  MoveL 497 to (87.59, -0.5, 58.1) mm, rotated rx 0 ry 90 rz 0 deg; joints [-13.797, -57.781, 117.086, 164.062, 60.282, -81.942]
  MoveL 498 to (93.3, -5.75, 58.1) mm, rotated rx 0 ry 90 rz 0 deg; joints [-13.739, -57.804, 116.577, 164.043, 59.762, -81.806]
  MoveL 499 to (99.9, -9.83, 58.1) mm, rotated rx 0 ry 90 rz 0 deg; joints [-13.673, -57.72, 116.001, 164.04, 59.279, -81.688]
  MoveL 500 to (107.03, -12.94, 58.1) mm, rotated rx 0 ry 90 rz 0 deg; joints [-13.603, -57.557, 115.386, 164.047, 58.834, -81.585]
  MoveL 501 to (114.36, -15.46, 58.1) mm, rotated rx 0 ry 90 rz 0 deg; joints [-13.531, -57.352, 114.755, 164.059, 58.415, -81.491]
  MoveL 502 to (121.65, -18.1, 58.1) mm, rotated rx 0 ry 90 rz 0 deg; joints [-13.46, -57.151, 114.125, 164.068, 57.991, -81.396]
  MoveL 503 to (126.38, -19.97, 58.1) mm, rotated rx 0 ry 90 rz 0 deg; joints [-13.414, -57.027, 113.713, 164.072, 57.707, -81.331]
  MoveL 504 to (131.09, -21.86, 58.1) mm, rotated rx 0 ry 90 rz 0 deg; joints [-13.369, -56.903, 113.3, 164.074, 57.422, -81.265]
  MoveL 505 to (135.76, -23.86, 58.1) mm, rotated rx 0 ry 90 rz 0 deg; joints [-13.325, -56.786, 112.889, 164.074, 57.133, -81.198]
  MoveL 506 to (140.36, -26.03, 58.1) mm, rotated rx 0 ry 90 rz 0 deg; joints [-13.281, -56.679, 112.48, 164.072, 56.837, -81.127]
  MoveL 507 to (145.03, -27.98, 58.1) mm, rotated rx 0 ry 90 rz 0 deg; joints [-13.237, -56.555, 112.066, 164.071, 56.55, -81.06]
  MoveL 508 to (150, -29.16, 58.1) mm, rotated rx 0 ry 90 rz 0 deg; joints [-13.191, -56.379, 111.633, 164.079, 56.296, -81.006]
  MoveL 509 to (150, -26.31, 58.1) mm, rotated rx 0 ry 90 rz 0 deg; joints [-13.191, -56.239, 111.66, 164.11, 56.456, -81.061]
  MoveL 510 to (146.2, -24.88, 58.1) mm, rotated rx 0 ry 90 rz 0 deg; joints [-13.226, -56.348, 111.996, 164.109, 56.681, -81.112]
  MoveL 511 to (142.73, -22.75, 58.1) mm, rotated rx 0 ry 90 rz 0 deg; joints [-13.259, -56.405, 112.31, 164.117, 56.932, -81.175]
  MoveL 512 to (139.28, -20.57, 58.1) mm, rotated rx 0 ry 90 rz 0 deg; joints [-13.291, -56.458, 112.622, 164.124, 57.187, -81.239]
  MoveL 513 to (135.74, -18.56, 58.1) mm, rotated rx 0 ry 90 rz 0 deg; joints [-13.325, -56.522, 112.938, 164.129, 57.434, -81.299]
  MoveL 514 to (132.21, -16.55, 58.1) mm, rotated rx 0 ry 90 rz 0 deg; joints [-13.358, -56.585, 113.253, 164.134, 57.682, -81.36]
  MoveL 515 to (127.82, -13.81, 58.1) mm, rotated rx 0 ry 90 rz 0 deg; joints [-13.4, -56.649, 113.645, 164.141, 58.004, -81.44]
  MoveL 516 to (123.5, -10.92, 58.1) mm, rotated rx 0 ry 90 rz 0 deg; joints [-13.442, -56.7, 114.031, 164.15, 58.332, -81.522]
  MoveL 517 to (119.33, -7.82, 58.1) mm, rotated rx 0 ry 90 rz 0 deg; joints [-13.482, -56.732, 114.405, 164.16, 58.666, -81.607]
  MoveL 518 to (115.6, -4.28, 58.1) mm, rotated rx 0 ry 90 rz 0 deg; joints [-13.518, -56.719, 114.744, 164.176, 59.011, -81.698]
  MoveL 519 to (112.62, 0, 58.1) mm, rotated rx 0 ry 90 rz 0 deg; joints [-13.548, -56.631, 115.024, 164.202, 59.369, -81.797]
  MoveL 520 to (-12.62, 0, 58.1) mm, rotated rx 0 ry 90 rz 0 deg; joints [-14.893, -62.159, 125.079, 163.369, 63.9, -82.514]
  MoveL 521 to (-15.6, -4.28, 58.1) mm, rotated rx 0 ry 90 rz 0 deg; joints [-14.928, -62.542, 125.276, 163.304, 63.726, -82.437]
  MoveL 522 to (-19.33, -7.82, 58.1) mm, rotated rx 0 ry 90 rz 0 deg; joints [-14.973, -62.916, 125.535, 163.239, 63.623, -82.379]
  MoveL 523 to (-23.5, -10.92, 58.1) mm, rotated rx 0 ry 90 rz 0 deg; joints [-15.023, -63.282, 125.831, 163.173, 63.561, -82.331]
  MoveL 524 to (-27.82, -13.81, 58.1) mm, rotated rx 0 ry 90 rz 0 deg; joints [-15.074, -63.645, 126.138, 163.108, 63.515, -82.287]
  MoveL 525 to (-32.2, -16.55, 58.1) mm, rotated rx 0 ry 90 rz 0 deg; joints [-15.128, -64.002, 126.45, 163.043, 63.478, -82.246]
  MoveL 526 to (-35.74, -18.56, 58.1) mm, rotated rx 0 ry 90 rz 0 deg; joints [-15.171, -64.279, 126.702, 162.991, 63.461, -82.217]
  MoveL 527 to (-39.28, -20.57, 58.1) mm, rotated rx 0 ry 90 rz 0 deg; joints [-15.214, -64.557, 126.953, 162.939, 63.442, -82.187]
  MoveL 528 to (-42.73, -22.75, 58.1) mm, rotated rx 0 ry 90 rz 0 deg; joints [-15.257, -64.841, 127.196, 162.886, 63.407, -82.152]
  MoveL 529 to (-46.2, -24.88, 58.1) mm, rotated rx 0 ry 90 rz 0 deg; joints [-15.3, -65.125, 127.439, 162.833, 63.375, -82.118]
  MoveL 530 to (-50, -26.31, 58.1) mm, rotated rx 0 ry 90 rz 0 deg; joints [-15.347, -65.381, 127.714, 162.783, 63.399, -82.1]
  MoveL 531 to (-50, -26.31, 103.1) mm, rotated rx 0 ry 90 rz 0 deg; joints [-17.375, -64.79, 126.71, 160.473, 63.306, -80.948]
  Sollgeschwindigkeit (200.0 mm/s)
  MoveL 532 to (-42.49, -26.16, 103.1) mm, rotated rx 0 ry 90 rz 0 deg; joints [-17.271, -64.448, 126.142, 160.55, 63.077, -80.915]
  MoveL 533 to (-34.99, -26.02, 103.1) mm, rotated rx 0 ry 90 rz 0 deg; joints [-17.168, -64.106, 125.572, 160.625, 62.845, -80.882]
  MoveL 534 to (-27.48, -25.87, 103.1) mm, rotated rx 0 ry 90 rz 0 deg; joints [-17.066, -63.763, 124.999, 160.699, 62.612, -80.848]
  MoveL 535 to (-19.97, -25.73, 103.1) mm, rotated rx 0 ry 90 rz 0 deg; joints [-16.966, -63.42, 124.425, 160.771, 62.377, -80.814]
  MoveL 536 to (-12.46, -25.58, 103.1) mm, rotated rx 0 ry 90 rz 0 deg; joints [-16.866, -63.077, 123.848, 160.842, 62.141, -80.778]
  MoveL 537 to (-4.96, -25.43, 103.1) mm, rotated rx 0 ry 90 rz 0 deg; joints [-16.768, -62.734, 123.268, 160.911, 61.902, -80.742]
  MoveL 538 to (2.55, -25.29, 103.1) mm, rotated rx 0 ry 90 rz 0 deg; joints [-16.671, -62.39, 122.687, 160.978, 61.661, -80.706]
  MoveL 539 to (10.05, -25.14, 103.1) mm, rotated rx 0 ry 90 rz 0 deg; joints [-16.575, -62.046, 122.103, 161.043, 61.419, -80.668]
  MoveL 540 to (17.56, -25, 103.1) mm, rotated rx 0 ry 90 rz 0 deg; joints [-16.48, -61.701, 121.516, 161.107, 61.175, -80.63]
  MoveL 541 to (25.07, -24.85, 103.1) mm, rotated rx 0 ry 90 rz 0 deg; joints [-16.386, -61.356, 120.927, 161.17, 60.929, -80.592]
  MoveL 542 to (32.58, -24.71, 103.1) mm, rotated rx 0 ry 90 rz 0 deg; joints [-16.293, -61.011, 120.336, 161.231, 60.681, -80.552]
  MoveL 543 to (40.08, -24.56, 103.1) mm, rotated rx 0 ry 90 rz 0 deg; joints [-16.201, -60.665, 119.742, 161.29, 60.431, -80.512]
  Sollgeschwindigkeit (50.0 mm/s)
  MoveL 544 to (40.08, -24.56, 58.1) mm, rotated rx 0 ry 90 rz 0 deg; joints [-14.296, -61.22, 120.719, 163.524, 60.538, -81.724]
  MoveL 545 to (36.66, -28.17, 58.1) mm, rotated rx 0 ry 90 rz 0 deg; joints [-14.334, -61.573, 120.955, 163.463, 60.432, -81.665]
  MoveL 546 to (36.08, -29.02, 58.1) mm, rotated rx 0 ry 90 rz 0 deg; joints [-14.34, -61.646, 120.993, 163.45, 60.399, -81.65]
  MoveL 547 to (35.49, -29.88, 58.1) mm, rotated rx 0 ry 90 rz 0 deg; joints [-14.346, -61.72, 121.031, 163.437, 60.366, -81.634]
  MoveL 548 to (34.9, -30.69, 58.08) mm, rotated rx 90 ry 86.96 rz 90 deg; joints [-14.257, -62.836, 120.907, 163.332, 59.164, -84.313]
  MoveL 549 to (34.32, -31.5, 58.01) mm, rotated rx 90 ry 83.41 rz 90 deg; joints [-14.096, -64.109, 120.741, 163.266, 57.761, -87.482]
  MoveL 550 to (33.73, -32.31, 57.9) mm, rotated rx 90 ry 79.85 rz 90 deg; joints [-13.873, -65.357, 120.562, 163.261, 56.359, -90.69]
  MoveL 551 to (33.17, -33.03, 57.74) mm, rotated rx 90 ry 76.63 rz 90 deg; joints [-13.62, -66.464, 120.392, 163.313, 55.094, -93.64]
  MoveL 552 to (32.6, -33.74, 57.55) mm, rotated rx 90 ry 73.4 rz 90 deg; joints [-13.318, -67.543, 120.214, 163.421, 53.837, -96.635]
  MoveL 553 to (32.04, -34.44, 57.32) mm, rotated rx 90 ry 70.18 rz 90 deg; joints [-12.968, -68.591, 120.028, 163.59, 52.593, -99.681]
  MoveL 554 to (31.48, -35.13, 57.05) mm, rotated rx 90 ry 66.95 rz 90 deg; joints [-12.57, -69.605, 119.836, 163.822, 51.364, -102.781]
  MoveL 555 to (30.63, -35.95, 56.67) mm, rotated rx 90 ry 63.01 rz 90 deg; joints [-12.022, -70.803, 119.607, 164.198, 49.895, -106.656]
  MoveL 556 to (29.79, -36.73, 56.24) mm, rotated rx 90 ry 59.07 rz 90 deg; joints [-11.405, -71.942, 119.374, 164.681, 48.463, -110.633]
  MoveL 557 to (28.94, -37.49, 55.75) mm, rotated rx 90 ry 55.13 rz 90 deg; joints [-10.723, -73.018, 119.14, 165.281, 47.076, -114.724]
  MoveL 558 to (28.04, -38.22, 55.2) mm, rotated rx 90 ry 51.13 rz 90 deg; joints [-9.964, -74.045, 118.907, 166.015, 45.723, -119.006]
  MoveL 559 to (27.13, -38.91, 54.6) mm, rotated rx 90 ry 47.13 rz 90 deg; joints [-9.143, -74.999, 118.678, 166.882, 44.436, -123.425]
  MoveL 560 to (26.62, -39.4, 54.13) mm, rotated rx 90 ry 44.19 rz 90 deg; joints [-8.5, -75.643, 118.503, 167.608, 43.534, -126.764]
  MoveL 561 to (26.11, -39.85, 53.64) mm, rotated rx 90 ry 41.24 rz 90 deg; joints [-7.827, -76.243, 118.333, 168.411, 42.677, -130.182]
  MoveL 562 to (25.61, -40.28, 53.12) mm, rotated rx 90 ry 38.3 rz 90 deg; joints [-7.124, -76.8, 118.17, 169.291, 41.869, -133.682]
  MoveL 563 to (25.48, -40.77, 52.46) mm, rotated rx 90 ry 34.73 rz 90 deg; joints [-6.232, -77.386, 117.944, 170.466, 40.951, -138.045]
  MoveL 564 to (25.37, -41.21, 51.78) mm, rotated rx 90 ry 31.15 rz 90 deg; joints [-5.304, -77.904, 117.731, 171.753, 40.121, -142.525]
  MoveL 565 to (25.25, -41.61, 51.06) mm, rotated rx 90 ry 27.57 rz 90 deg; joints [-4.344, -78.351, 117.534, 173.144, 39.385, -147.116]
  MoveL 566 to (25.45, -41.88, 50.53) mm, rotated rx 90 ry 24.95 rz 90 deg; joints [-3.621, -78.616, 117.379, 174.228, 38.905, -150.548]
  MoveL 567 to (25.65, -42.12, 49.98) mm, rotated rx 90 ry 22.33 rz 90 deg; joints [-2.886, -78.842, 117.233, 175.359, 38.482, -154.03]
  MoveL 568 to (26.42, -42.43, 49.12) mm, rotated rx 90 ry 18.35 rz 90 deg; joints [-1.747, -79.083, 116.996, 177.159, 37.948, -159.407]
  MoveL 569 to (27.19, -42.54, 48.79) mm, rotated rx 90 ry 16.83 rz 90 deg; joints [-1.304, -79.122, 116.877, 177.871, 37.774, -161.491]
  MoveL 570 to (27.95, -42.64, 48.46) mm, rotated rx 90 ry 15.3 rz 90 deg; joints [-0.86, -79.147, 116.761, 178.592, 37.622, -163.585]
  MoveL 571 to (28.72, -42.72, 48.12) mm, rotated rx 90 ry 13.77 rz 90 deg; joints [-0.413, -79.159, 116.649, 179.321, 37.492, -165.687]
  MoveL 572 to (29.56, -42.79, 47.84) mm, rotated rx 90 ry 12.53 rz 90 deg; joints [-0.048, -79.145, 116.544, 179.921, 37.398, -167.409]
  MoveL 573 to (30.4, -42.85, 47.56) mm, rotated rx 90 ry 11.28 rz 90 deg; joints [0.318, -79.123, 116.442, -179.476, 37.32, -169.135]
  MoveL 574 to (31.24, -42.9, 47.28) mm, rotated rx 90 ry 10.04 rz 90 deg; joints [0.684, -79.092, 116.342, -178.87, 37.256, -170.862]
  MoveL 575 to (31.96, -42.97, 46.87) mm, rotated rx 90 ry 8.2 rz 90 deg; joints [1.225, -79.061, 116.239, -177.974, 37.195, -173.413]
  MoveL 576 to (32.69, -43.02, 46.45) mm, rotated rx 90 ry 6.37 rz 90 deg; joints [1.765, -79.012, 116.143, -177.078, 37.167, -175.965]
  MoveL 577 to (33.42, -43.06, 46.03) mm, rotated rx 90 ry 4.53 rz 90 deg; joints [2.305, -78.943, 116.052, -176.183, 37.17, -178.514]
  MoveL 578 to (34.18, -43.09, 45.39) mm, rotated rx 90 ry 1.71 rz 90 deg; joints [3.132, -78.823, 115.951, -174.82, 37.241, 177.584]
  MoveL 579 to (34.94, -43.1, 44.73) mm, rotated rx 90 ry 0 rz 90 deg; joints [3.644, -78.708, 115.873, -173.982, 37.317, 175.208]
  MoveL 580 to (35.7, -43.1, 44.06) mm, rotated rx 90 ry 0 rz 90 deg; joints [3.672, -78.658, 115.812, -173.934, 37.308, 175.169]
  MoveL 581 to (37.13, -43.1, 42.71) mm, rotated rx 90 ry 0 rz 90 deg; joints [3.729, -78.564, 115.695, -173.837, 37.292, 175.09]
  MoveL 582 to (38.7, -43.1, 41.89) mm, rotated rx 90 ry 0 rz 90 deg; joints [3.762, -78.463, 115.572, -173.78, 37.272, 175.043]
  MoveL 583 to (40.05, -43.1, 41.81) mm, rotated rx 90 ry 0 rz 90 deg; joints [3.762, -78.378, 115.468, -173.778, 37.252, 175.04]
  MoveL 584 to (41.5, -43.1, 42.11) mm, rotated rx 90 ry 0 rz 90 deg; joints [3.744, -78.29, 115.359, -173.805, 37.231, 175.06]
  MoveL 585 to (45.39, -43.1, 43.71) mm, rotated rx 90 ry 0 rz 90 deg; joints [3.66, -78.055, 115.069, -173.934, 37.169, 175.16]
  MoveL 586 to (47.73, -43.1, 44.54) mm, rotated rx 90 ry 0 rz 90 deg; joints [3.616, -77.913, 114.892, -174.003, 37.131, 175.212]
  MoveL 587 to (50.09, -43.1, 44.8) mm, rotated rx 90 ry 0 rz 90 deg; joints [3.598, -77.767, 114.712, -174.028, 37.095, 175.23]
  MoveL 588 to (53.81, -43.1, 44.03) mm, rotated rx 90 ry 0 rz 90 deg; joints [3.621, -77.534, 114.421, -173.981, 37.04, 175.189]
  MoveL 589 to (56.17, -43.1, 43.02) mm, rotated rx 90 ry 0 rz 90 deg; joints [3.66, -77.383, 114.234, -173.912, 37.006, 175.132]
  MoveL 590 to (58.51, -43.1, 42.11) mm, rotated rx 90 ry 0 rz 90 deg; joints [3.694, -77.235, 114.049, -173.85, 36.972, 175.08]
  MoveL 591 to (60.69, -43.1, 41.79) mm, rotated rx 90 ry 0 rz 90 deg; joints [3.702, -77.099, 113.877, -173.832, 36.938, 175.064]
  MoveL 592 to (62.64, -43.1, 42.54) mm, rotated rx 90 ry 0 rz 90 deg; joints [3.663, -76.981, 113.73, -173.893, 36.905, 175.11]
  MoveL 593 to (64.38, -43.1, 44.14) mm, rotated rx 90 ry 0 rz 90 deg; joints [3.587, -76.88, 113.602, -174.015, 36.872, 175.206]
  MoveL 594 to (65.25, -43.1, 44.93) mm, rotated rx 90 ry 0 rz 90 deg; joints [3.549, -76.829, 113.538, -174.076, 36.856, 175.254]
  MoveL 595 to (66.12, -43.08, 45.69) mm, rotated rx 90 ry 3.02 rz 90 deg; joints [2.68, -76.878, 113.508, -175.514, 36.714, 179.42]
  MoveL 596 to (66.83, -43.05, 46.15) mm, rotated rx 90 ry 5.01 rz 90 deg; joints [2.106, -76.874, 113.486, -176.471, 36.664, -177.819]
  MoveL 597 to (67.55, -43, 46.6) mm, rotated rx 90 ry 7.01 rz 90 deg; joints [1.533, -76.848, 113.471, -177.431, 36.65, -175.056]
  MoveL 598 to (68.26, -42.94, 47.05) mm, rotated rx 90 ry 9 rz 90 deg; joints [0.961, -76.8, 113.463, -178.391, 36.673, -172.291]
  MoveL 599 to (69.09, -42.89, 47.36) mm, rotated rx 90 ry 10.36 rz 90 deg; joints [0.571, -76.734, 113.434, -179.045, 36.704, -170.404]
  MoveL 600 to (69.93, -42.83, 47.66) mm, rotated rx 90 ry 11.72 rz 90 deg; joints [0.182, -76.657, 113.408, -179.695, 36.751, -168.52]
  MoveL 601 to (70.76, -42.76, 47.97) mm, rotated rx 90 ry 13.09 rz 90 deg; joints [-0.205, -76.57, 113.385, 179.658, 36.816, -166.639]
  MoveL 602 to (71.58, -42.68, 48.27) mm, rotated rx 90 ry 14.47 rz 90 deg; joints [-0.596, -76.473, 113.367, 179.007, 36.898, -164.738]
  MoveL 603 to (72.39, -42.6, 48.58) mm, rotated rx 90 ry 15.85 rz 90 deg; joints [-0.984, -76.366, 113.353, 178.364, 36.998, -162.844]
  MoveL 604 to (73.21, -42.51, 48.88) mm, rotated rx 90 ry 17.23 rz 90 deg; joints [-1.371, -76.248, 113.341, 177.728, 37.114, -160.958]
  MoveL 605 to (74.11, -42.25, 49.63) mm, rotated rx 90 ry 20.72 rz 90 deg; joints [-2.336, -75.977, 113.415, 176.162, 37.5, -156.237]
  MoveL 606 to (74.39, -42.04, 50.16) mm, rotated rx 90 ry 23.19 rz 90 deg; joints [-3.01, -75.767, 113.508, 175.09, 37.843, -152.928]
  MoveL 607 to (74.66, -41.81, 50.67) mm, rotated rx 90 ry 25.67 rz 90 deg; joints [-3.674, -75.524, 113.609, 174.057, 38.235, -149.659]
  MoveL 608 to (74.68, -41.51, 51.25) mm, rotated rx 90 ry 28.48 rz 90 deg; joints [-4.416, -75.226, 113.757, 172.933, 38.744, -145.993]
  MoveL 609 to (74.71, -41.19, 51.81) mm, rotated rx 90 ry 31.3 rz 90 deg; joints [-5.141, -74.885, 113.915, 171.869, 39.313, -142.39]
  MoveL 610 to (74.73, -40.84, 52.35) mm, rotated rx 90 ry 34.12 rz 90 deg; joints [-5.847, -74.503, 114.082, 170.868, 39.938, -138.854]
  MoveL 611 to (74.34, -40.35, 53.03) mm, rotated rx 90 ry 37.83 rz 90 deg; joints [-6.748, -73.962, 114.347, 169.651, 40.85, -134.301]
  MoveL 612 to (73.95, -39.8, 53.69) mm, rotated rx 90 ry 41.55 rz 90 deg; joints [-7.609, -73.352, 114.626, 168.551, 41.846, -129.873]
  MoveL 613 to (73.31, -39.3, 54.23) mm, rotated rx 90 ry 44.78 rz 90 deg; joints [-8.327, -72.782, 114.901, 167.689, 42.783, -126.115]
  MoveL 614 to (72.67, -38.76, 54.74) mm, rotated rx 90 ry 48.02 rz 90 deg; joints [-9.01, -72.161, 115.181, 166.916, 43.773, -122.452]
  MoveL 615 to (71.98, -38.23, 55.19) mm, rotated rx 90 ry 51.07 rz 90 deg; joints [-9.619, -71.538, 115.457, 166.269, 44.75, -119.09]
  MoveL 616 to (71.29, -37.68, 55.61) mm, rotated rx 90 ry 54.11 rz 90 deg; joints [-10.195, -70.872, 115.736, 165.698, 45.765, -115.806]
  MoveL 617 to (70.43, -36.92, 56.12) mm, rotated rx 90 ry 58.1 rz 90 deg; joints [-10.895, -69.937, 116.1, 165.058, 47.147, -111.615]
  MoveL 618 to (69.56, -36.13, 56.58) mm, rotated rx 90 ry 62.09 rz 90 deg; joints [-11.532, -68.935, 116.464, 164.537, 48.579, -107.543]
  MoveL 619 to (68.7, -35.31, 56.97) mm, rotated rx 90 ry 66.07 rz 90 deg; joints [-12.103, -67.872, 116.825, 164.127, 50.054, -103.58]
  MoveL 620 to (68.12, -34.62, 57.26) mm, rotated rx 90 ry 69.32 rz 90 deg; joints [-12.517, -66.955, 117.105, 163.871, 51.278, -100.423]
  MoveL 621 to (67.54, -33.92, 57.5) mm, rotated rx 90 ry 72.57 rz 90 deg; joints [-12.885, -66.002, 117.38, 163.68, 52.522, -97.325]
  MoveL 622 to (66.97, -33.21, 57.7) mm, rotated rx 90 ry 75.82 rz 90 deg; joints [-13.205, -65.016, 117.648, 163.551, 53.78, -94.281]
  MoveL 623 to (66.39, -32.48, 57.86) mm, rotated rx 90 ry 79.07 rz 90 deg; joints [-13.478, -64, 117.908, 163.48, 55.05, -91.284]
  MoveL 624 to (65.8, -31.67, 57.99) mm, rotated rx 90 ry 82.69 rz 90 deg; joints [-13.723, -62.836, 118.183, 163.466, 56.47, -88.001]
  MoveL 625 to (65.21, -30.85, 58.07) mm, rotated rx 90 ry 86.3 rz 90 deg; joints [-13.908, -61.643, 118.445, 163.515, 57.895, -84.763]
  MoveL 626 to (64.61, -30.02, 58.1) mm, rotated rx 90 ry 89.91 rz 90 deg; joints [-14.032, -60.424, 118.693, 163.625, 59.32, -81.561]
  MoveL 627 to (64.02, -29.15, 58.1) mm, rotated rx 0 ry 90 rz 0 deg; joints [-14.04, -60.376, 118.754, 163.633, 59.426, -81.504]
  MoveL 628 to (63.42, -28.29, 58.1) mm, rotated rx 0 ry 90 rz 0 deg; joints [-14.047, -60.357, 118.81, 163.639, 59.5, -81.525]
  MoveL 629 to (59.97, -24.61, 58.1) mm, rotated rx 0 ry 90 rz 0 deg; joints [-14.083, -60.318, 119.125, 163.655, 59.844, -81.619]
  MoveL 630 to (55.88, -21.25, 58.1) mm, rotated rx 0 ry 90 rz 0 deg; joints [-14.126, -60.323, 119.486, 163.664, 60.192, -81.71]
  MoveL 631 to (53.52, -19.72, 58.1) mm, rotated rx 0 ry 90 rz 0 deg; joints [-14.152, -60.348, 119.69, 163.664, 60.368, -81.754]
  MoveL 632 to (50.78, -19.09, 58.1) mm, rotated rx 0 ry 90 rz 0 deg; joints [-14.181, -60.437, 119.915, 163.652, 60.502, -81.782]
  MoveL 633 to (47.22, -19.46, 58.1) mm, rotated rx 0 ry 90 rz 0 deg; joints [-14.219, -60.618, 120.197, 163.625, 60.605, -81.793]
  MoveL 634 to (44.12, -21.25, 58.1) mm, rotated rx 0 ry 90 rz 0 deg; joints [-14.253, -60.856, 120.428, 163.586, 60.603, -81.772]
  MoveL 635 to (44.07, -28.84, 58.1) mm, rotated rx 0 ry 90 rz 0 deg; joints [-14.253, -61.272, 120.358, 163.507, 60.137, -81.613]
  MoveL 636 to (43.49, -29.77, 58.1) mm, rotated rx 0 ry 90 rz 0 deg; joints [-14.259, -61.348, 120.395, 163.493, 60.1, -81.597]
  MoveL 637 to (42.91, -30.65, 58.08) mm, rotated rx 90 ry 87.14 rz 90 deg; joints [-14.177, -62.399, 120.28, 163.392, 58.97, -84.12]
  MoveL 638 to (42.34, -31.53, 58.01) mm, rotated rx 90 ry 83.3 rz 90 deg; joints [-14.004, -63.761, 120.098, 163.32, 57.465, -87.545]
  MoveL 639 to (41.88, -32.37, 57.88) mm, rotated rx 90 ry 79.6 rz 90 deg; joints [-13.769, -65.04, 119.901, 163.319, 56.012, -90.891]
  MoveL 640 to (41.43, -33.19, 57.71) mm, rotated rx 90 ry 75.9 rz 90 deg; joints [-13.47, -66.286, 119.69, 163.389, 54.566, -94.29]
  MoveL 641 to (40.98, -34.01, 57.47) mm, rotated rx 90 ry 72.2 rz 90 deg; joints [-13.107, -67.494, 119.469, 163.534, 53.133, -97.749]
  MoveL 642 to (40.72, -34.71, 57.23) mm, rotated rx 90 ry 68.95 rz 90 deg; joints [-12.734, -68.513, 119.256, 163.73, 51.886, -100.842]
  MoveL 643 to (40.45, -35.39, 56.94) mm, rotated rx 90 ry 65.7 rz 90 deg; joints [-12.315, -69.496, 119.038, 163.991, 50.657, -103.995]
  MoveL 644 to (40.19, -36.06, 56.61) mm, rotated rx 90 ry 62.45 rz 90 deg; joints [-11.848, -70.441, 118.816, 164.323, 49.451, -107.214]
  MoveL 645 to (40.09, -36.77, 56.21) mm, rotated rx 90 ry 58.87 rz 90 deg; joints [-11.281, -71.423, 118.555, 164.775, 48.151, -110.837]
  MoveL 646 to (39.98, -37.46, 55.77) mm, rotated rx 90 ry 55.3 rz 90 deg; joints [-10.661, -72.352, 118.293, 165.321, 46.89, -114.554]
  MoveL 647 to (39.87, -38.12, 55.28) mm, rotated rx 90 ry 51.72 rz 90 deg; joints [-9.989, -73.226, 118.033, 165.968, 45.675, -118.371]
  MoveL 648 to (40.01, -38.71, 54.79) mm, rotated rx 90 ry 48.34 rz 90 deg; joints [-9.305, -73.986, 117.771, 166.678, 44.565, -122.088]
  MoveL 649 to (40.14, -39.27, 54.26) mm, rotated rx 90 ry 44.95 rz 90 deg; joints [-8.579, -74.692, 117.514, 167.486, 43.509, -125.905]
  MoveL 650 to (40.28, -39.8, 53.69) mm, rotated rx 90 ry 41.56 rz 90 deg; joints [-7.814, -75.342, 117.264, 168.393, 42.511, -129.828]
  MoveL 651 to (41.08, -40.38, 52.98) mm, rotated rx 90 ry 37.55 rz 90 deg; joints [-6.855, -75.998, 116.93, 169.602, 41.402, -134.613]
  MoveL 652 to (41.87, -40.92, 52.24) mm, rotated rx 90 ry 33.54 rz 90 deg; joints [-5.851, -76.569, 116.611, 170.95, 40.396, -139.547]
  MoveL 653 to (42.67, -41.4, 51.45) mm, rotated rx 90 ry 29.52 rz 90 deg; joints [-4.804, -77.054, 116.31, 172.434, 39.502, -144.625]
  MoveL 654 to (43.46, -41.59, 51.1) mm, rotated rx 90 ry 27.73 rz 90 deg; joints [-4.324, -77.215, 116.149, 173.139, 39.135, -146.934]
  MoveL 655 to (44.24, -41.78, 50.73) mm, rotated rx 90 ry 25.94 rz 90 deg; joints [-3.838, -77.359, 115.992, 173.868, 38.794, -149.27]
  MoveL 656 to (45.03, -41.95, 50.36) mm, rotated rx 90 ry 24.15 rz 90 deg; joints [-3.345, -77.485, 115.84, 174.619, 38.478, -151.631]
  MoveL 657 to (45.82, -42.12, 49.98) mm, rotated rx 90 ry 22.36 rz 90 deg; joints [-2.848, -77.593, 115.692, 175.391, 38.189, -154.014]
  MoveL 658 to (46.7, -42.18, 49.83) mm, rotated rx 90 ry 21.64 rz 90 deg; joints [-2.645, -77.596, 115.59, 175.708, 38.072, -154.978]
  MoveL 659 to (47.59, -42.24, 49.68) mm, rotated rx 90 ry 20.92 rz 90 deg; joints [-2.442, -77.596, 115.489, 176.028, 37.959, -155.946]
  MoveL 660 to (48.48, -42.29, 49.52) mm, rotated rx 90 ry 20.2 rz 90 deg; joints [-2.238, -77.593, 115.388, 176.351, 37.851, -156.916]
  MoveL 661 to (49.36, -42.35, 49.37) mm, rotated rx 90 ry 19.48 rz 90 deg; joints [-2.034, -77.588, 115.289, 176.676, 37.748, -157.89]
  MoveL 662 to (50.21, -42.32, 49.46) mm, rotated rx 90 ry 19.89 rz 90 deg; joints [-2.148, -77.508, 115.241, 176.493, 37.785, -157.336]
  MoveL 663 to (51.06, -42.29, 49.55) mm, rotated rx 90 ry 20.3 rz 90 deg; joints [-2.262, -77.427, 115.193, 176.31, 37.824, -156.783]
  MoveL 664 to (51.9, -42.25, 49.63) mm, rotated rx 90 ry 20.71 rz 90 deg; joints [-2.375, -77.345, 115.146, 176.129, 37.864, -156.231]
  MoveL 665 to (52.75, -42.22, 49.72) mm, rotated rx 90 ry 21.12 rz 90 deg; joints [-2.487, -77.263, 115.099, 175.949, 37.906, -155.682]
  MoveL 666 to (53.6, -42.19, 49.81) mm, rotated rx 90 ry 21.53 rz 90 deg; joints [-2.6, -77.179, 115.052, 175.77, 37.949, -155.132]
  MoveL 667 to (54.54, -42.01, 50.24) mm, rotated rx 90 ry 23.57 rz 90 deg; joints [-3.161, -76.952, 115.076, 174.888, 38.234, -152.411]
  MoveL 668 to (55.49, -41.81, 50.66) mm, rotated rx 90 ry 25.61 rz 90 deg; joints [-3.714, -76.703, 115.105, 174.034, 38.554, -149.717]
  MoveL 669 to (56.43, -41.6, 51.08) mm, rotated rx 90 ry 27.65 rz 90 deg; joints [-4.258, -76.431, 115.14, 173.21, 38.906, -147.055]
  MoveL 670 to (57.37, -41.38, 51.49) mm, rotated rx 90 ry 29.69 rz 90 deg; joints [-4.793, -76.137, 115.18, 172.418, 39.29, -144.427]
  MoveL 671 to (58.13, -41.03, 52.07) mm, rotated rx 90 ry 32.65 rz 90 deg; joints [-5.552, -75.71, 115.295, 171.327, 39.91, -140.677]
  MoveL 672 to (58.88, -40.65, 52.63) mm, rotated rx 90 ry 35.61 rz 90 deg; joints [-6.288, -75.236, 115.42, 170.309, 40.59, -137.004]
  MoveL 673 to (59.36, -40.15, 53.28) mm, rotated rx 90 ry 39.22 rz 90 deg; joints [-7.155, -74.625, 115.618, 169.166, 41.504, -132.625]
  MoveL 674 to (59.83, -39.61, 53.91) mm, rotated rx 90 ry 42.83 rz 90 deg; joints [-7.982, -73.948, 115.827, 168.137, 42.495, -128.365]
  MoveL 675 to (59.93, -39.14, 54.38) mm, rotated rx 90 ry 45.74 rz 90 deg; joints [-8.619, -73.373, 116.025, 167.39, 43.349, -125.02]
  MoveL 676 to (60.03, -38.66, 54.83) mm, rotated rx 90 ry 48.65 rz 90 deg; joints [-9.226, -72.759, 116.227, 166.716, 44.245, -121.752]
  MoveL 677 to (60.13, -38.15, 55.26) mm, rotated rx 90 ry 51.56 rz 90 deg; joints [-9.802, -72.105, 116.432, 166.112, 45.178, -118.556]
  MoveL 678 to (60.05, -37.59, 55.68) mm, rotated rx 90 ry 54.61 rz 90 deg; joints [-10.374, -71.388, 116.665, 165.552, 46.197, -115.279]
  MoveL 679 to (59.98, -37.01, 56.07) mm, rotated rx 90 ry 57.66 rz 90 deg; joints [-10.909, -70.631, 116.898, 165.066, 47.249, -112.078]
  MoveL 680 to (59.9, -36.41, 56.43) mm, rotated rx 90 ry 60.71 rz 90 deg; joints [-11.406, -69.836, 117.132, 164.649, 48.332, -108.945]
  MoveL 681 to (59.62, -35.65, 56.82) mm, rotated rx 90 ry 64.44 rz 90 deg; joints [-11.962, -68.826, 117.43, 164.229, 49.692, -105.211]
  MoveL 682 to (59.34, -34.88, 57.16) mm, rotated rx 90 ry 68.16 rz 90 deg; joints [-12.458, -67.764, 117.724, 163.903, 51.084, -101.567]
  MoveL 683 to (59.05, -34.07, 57.45) mm, rotated rx 90 ry 71.88 rz 90 deg; joints [-12.894, -66.655, 118.011, 163.665, 52.502, -98.003]
  MoveL 684 to (58.63, -33.3, 57.68) mm, rotated rx 90 ry 75.43 rz 90 deg; joints [-13.253, -65.565, 118.29, 163.513, 53.878, -94.673]
  MoveL 685 to (58.2, -32.51, 57.86) mm, rotated rx 90 ry 78.98 rz 90 deg; joints [-13.554, -64.438, 118.56, 163.431, 55.268, -91.4]
  MoveL 686 to (57.77, -31.7, 57.99) mm, rotated rx 90 ry 82.53 rz 90 deg; joints [-13.797, -63.279, 118.819, 163.415, 56.667, -88.178]
  MoveL 687 to (57.22, -30.86, 58.07) mm, rotated rx 90 ry 86.22 rz 90 deg; joints [-13.989, -62.045, 119.083, 163.463, 58.133, -84.866]
  MoveL 688 to (56.68, -30.02, 58.1) mm, rotated rx 90 ry 89.92 rz 90 deg; joints [-14.116, -60.784, 119.333, 163.575, 59.601, -81.593]
  MoveL 689 to (56.13, -29.13, 58.1) mm, rotated rx 0 ry 90 rz 0 deg; joints [-14.124, -60.736, 119.389, 163.584, 59.703, -81.546]
  MoveL 690 to (53.89, -27.09, 58.1) mm, rotated rx 0 ry 90 rz 0 deg; joints [-14.148, -60.729, 119.59, 163.59, 59.905, -81.6]
  MoveL 691 to (50.99, -26.34, 58.1) mm, rotated rx 0 ry 90 rz 0 deg; joints [-14.179, -60.82, 119.829, 163.579, 60.052, -81.63]
  MoveL 692 to (48.41, -26.38, 58.1) mm, rotated rx 0 ry 90 rz 0 deg; joints [-14.206, -60.94, 120.036, 163.562, 60.139, -81.643]
  MoveL 693 to (45.99, -27.16, 58.1) mm, rotated rx 0 ry 90 rz 0 deg; joints [-14.232, -61.093, 120.222, 163.537, 60.174, -81.639]
  MoveL 694 to (44.07, -28.84, 58.1) mm, rotated rx 0 ry 90 rz 0 deg; joints [-14.253, -61.272, 120.358, 163.507, 60.137, -81.613]
  MoveL 695 to (44.07, -28.84, 103.1) mm, rotated rx 0 ry 90 rz 0 deg; joints [-16.152, -60.715, 119.383, 161.27, 60.035, -80.388]
  Sollgeschwindigkeit (200.0 mm/s)
  MoveL 696 to (47.12, -37.25, 102.65) mm, rotated rx 90 ry 82.83 rz 90 deg; joints [-15.812, -63.405, 118.665, 160.985, 56.749, -86.47]
  MoveL 697 to (50.18, -47.77, 100.32) mm, rotated rx 90 ry 72.19 rz 90 deg; joints [-14.835, -67.11, 117.621, 161.058, 52.068, -95.897]
  MoveL 698 to (53.23, -57.68, 96.08) mm, rotated rx 90 ry 61.55 rz 90 deg; joints [-13.293, -70.401, 116.489, 161.844, 47.548, -105.967]
  MoveL 699 to (56.28, -66.63, 90.1) mm, rotated rx 90 ry 50.91 rz 90 deg; joints [-11.222, -73.187, 115.329, 163.527, 43.338, -116.95]
  MoveL 700 to (59.34, -74.33, 82.56) mm, rotated rx 90 ry 40.27 rz 90 deg; joints [-8.679, -75.395, 114.207, 166.312, 39.62, -129.1]
  MoveL 701 to (62.39, -80.5, 73.73) mm, rotated rx 90 ry 29.64 rz 90 deg; joints [-5.745, -76.97, 113.188, 170.336, 36.609, -142.581]
  MoveL 702 to (65.44, -84.94, 63.91) mm, rotated rx 90 ry 19 rz 90 deg; joints [-2.526, -77.877, 112.33, 175.542, 34.534, -157.329]
  MoveL 703 to (68.49, -87.48, 53.45) mm, rotated rx 90 ry 8.36 rz 90 deg; joints [0.854, -78.1, 111.677, -178.456, 33.587, -172.93]
  MoveL 704 to (71.55, -88.1, 44.24) mm, rotated rx 90 ry 0 rz 90 deg; joints [3.563, -77.75, 111.269, -173.567, 33.685, 174.64]
  MoveL 705 to (74.6, -88.1, 40.69) mm, rotated rx 90 ry 0 rz 90 deg; joints [3.711, -77.544, 111.013, -173.293, 33.65, 174.409]
  MoveL 706 to (77.65, -88.1, 37.15) mm, rotated rx 90 ry 0 rz 90 deg; joints [3.858, -77.337, 110.757, -173.02, 33.615, 174.178]
  MoveL 707 to (80.71, -88.1, 33.6) mm, rotated rx 90 ry 0 rz 90 deg; joints [4.004, -77.13, 110.499, -172.747, 33.58, 173.947]
  MoveL 708 to (83.76, -88.1, 30.05) mm, rotated rx 90 ry 0 rz 90 deg; joints [4.15, -76.923, 110.239, -172.475, 33.544, 173.717]
  MoveL 709 to (86.81, -88.1, 26.51) mm, rotated rx 90 ry 0 rz 90 deg; joints [4.295, -76.715, 109.979, -172.203, 33.508, 173.487]
  MoveL 710 to (89.87, -88.1, 22.96) mm, rotated rx 90 ry 0 rz 90 deg; joints [4.439, -76.507, 109.717, -171.933, 33.472, 173.257]
  MoveL 711 to (92.92, -88.1, 19.42) mm, rotated rx 90 ry 0 rz 90 deg; joints [4.583, -76.298, 109.454, -171.662, 33.435, 173.027]
  MoveL 712 to (95.97, -88.1, 15.87) mm, rotated rx 90 ry 0 rz 90 deg; joints [4.726, -76.089, 109.189, -171.393, 33.398, 172.798]
  MoveL 713 to (99.03, -87.53, 6.88) mm, rotated rx 90 ry -8.03 rz 90 deg; joints [7.22, -75.287, 108.808, -167.08, 34.201, 161.226]
  MoveL 714 to (102.08, -85.04, -3.6) mm, rotated rx 90 ry -18.67 rz 90 deg; joints [10.302, -73.748, 108.585, -162.348, 36.142, 146.918]
  MoveL 715 to (105.13, -80.66, -13.44) mm, rotated rx 90 ry -29.31 rz 90 deg; joints [13.082, -71.635, 108.559, -158.853, 38.86, 133.93]
  MoveL 716 to (108.18, -74.54, -22.3) mm, rotated rx 90 ry -39.95 rz 90 deg; joints [15.471, -69.007, 108.695, -156.567, 42.127, 122.233]
  MoveL 717 to (111.24, -66.89, -29.89) mm, rotated rx 90 ry -50.59 rz 90 deg; joints [17.405, -65.936, 108.944, -155.317, 45.751, 111.633]
  MoveL 718 to (114.29, -57.97, -35.93) mm, rotated rx 90 ry -61.22 rz 90 deg; joints [18.843, -62.503, 109.259, -154.898, 49.58, 101.878]
  MoveL 719 to (117.34, -48.09, -40.21) mm, rotated rx 90 ry -71.86 rz 90 deg; joints [19.758, -58.798, 109.594, -155.13, 53.497, 92.72]
  MoveL 720 to (120.4, -37.58, -42.6) mm, rotated rx 90 ry -82.5 rz 90 deg; joints [20.139, -54.923, 109.912, -155.88, 57.408, 83.939]
  MoveL 721 to (123.45, -28.95, -43.1) mm, rotated rx 0 ry -90 rz 180 deg; joints [20.071, -52.056, 110.04, -156.688, 60.135, 77.889]
  MoveL 722 to (126.5, -25.41, -43.1) mm, rotated rx 0 ry -90 rz 180 deg; joints [20.029, -51.745, 109.8, -156.751, 60.191, 77.945]
  MoveL 723 to (129.56, -21.86, -43.1) mm, rotated rx 0 ry -90 rz 180 deg; joints [19.988, -51.433, 109.558, -156.814, 60.247, 78]
  MoveL 724 to (132.61, -18.31, -43.1) mm, rotated rx 0 ry -90 rz 180 deg; joints [19.946, -51.122, 109.314, -156.876, 60.3, 78.054]
  MoveL 725 to (135.66, -14.77, -43.1) mm, rotated rx 0 ry -90 rz 180 deg; joints [19.905, -50.811, 109.069, -156.937, 60.353, 78.107]
  MoveL 726 to (138.72, -11.22, -43.1) mm, rotated rx 0 ry -90 rz 180 deg; joints [19.864, -50.5, 108.823, -156.998, 60.403, 78.158]
  MoveL 727 to (141.77, -7.67, -43.1) mm, rotated rx 0 ry -90 rz 180 deg; joints [19.822, -50.189, 108.574, -157.058, 60.452, 78.209]
  MoveL 728 to (144.82, -4.13, -43.1) mm, rotated rx 0 ry -90 rz 180 deg; joints [19.782, -49.878, 108.324, -157.117, 60.5, 78.259]
  Sollgeschwindigkeit (50.0 mm/s)
  MoveL 729 to (144.82, -4.13, 1.9) mm, rotated rx 0 ry -90 rz 180 deg; joints [18.092, -50.536, 109.633, -159.156, 60.778, 79.47]
  MoveL 730 to (139.38, -5.04, 1.9) mm, rotated rx 0 ry -90 rz 180 deg; joints [18.159, -50.814, 110.091, -159.116, 60.958, 79.507]
  MoveL 731 to (133.91, -5.84, 1.9) mm, rotated rx 0 ry -90 rz 180 deg; joints [18.228, -51.088, 110.55, -159.075, 61.144, 79.545]
  MoveL 732 to (128.63, -7.16, 1.9) mm, rotated rx 0 ry -90 rz 180 deg; joints [18.294, -51.38, 110.99, -159.03, 61.294, 79.569]
  MoveL 733 to (123.52, -9.64, 1.9) mm, rotated rx 0 ry -90 rz 180 deg; joints [18.359, -51.726, 111.411, -158.972, 61.376, 79.565]
  MoveL 734 to (118.88, -13.11, 1.9) mm, rotated rx 0 ry -90 rz 180 deg; joints [18.419, -52.103, 111.788, -158.905, 61.386, 79.533]
  MoveL 735 to (114.74, -17.2, 1.9) mm, rotated rx 0 ry -90 rz 180 deg; joints [18.472, -52.494, 112.119, -158.834, 61.34, 79.48]
  MoveL 736 to (112.95, -19.92, 1.9) mm, rotated rx 0 ry -90 rz 180 deg; joints [18.495, -52.712, 112.258, -158.792, 61.271, 79.435]
  MoveL 737 to (112.03, -23.12, 1.9) mm, rotated rx 0 ry -90 rz 180 deg; joints [18.507, -52.919, 112.323, -158.75, 61.141, 79.37]
  MoveL 738 to (112.11, -25.32, 1.9) mm, rotated rx 0 ry -90 rz 180 deg; joints [18.506, -53.031, 112.308, -158.726, 61.022, 79.318]
  MoveL 739 to (112.9, -27.3, 1.9) mm, rotated rx 0 ry -90 rz 180 deg; joints [18.496, -53.101, 112.234, -158.709, 60.886, 79.264]
  MoveL 740 to (114.27, -29, 1.9) mm, rotated rx 0 ry -90 rz 180 deg; joints [18.478, -53.13, 112.113, -158.698, 60.743, 79.211]
  MoveL 741 to (115.1, -29.83, 1.9) mm, rotated rx 0 ry -90 rz 180 deg; joints [18.467, -53.138, 112.041, -158.694, 60.667, 79.183]
  MoveL 742 to (115.92, -30.62, 1.92) mm, rotated rx 90 ry -87.28 rz 90 deg; joints [18.5, -53.995, 111.852, -158.438, 59.699, 81.439]
  MoveL 743 to (116.74, -31.41, 1.98) mm, rotated rx 90 ry -83.84 rz 90 deg; joints [18.498, -55.076, 111.627, -158.151, 58.485, 84.318]
  MoveL 744 to (117.57, -32.18, 2.08) mm, rotated rx 90 ry -80.4 rz 90 deg; joints [18.444, -56.151, 111.4, -157.907, 57.266, 87.216]
  MoveL 745 to (118.39, -32.96, 2.24) mm, rotated rx 90 ry -76.96 rz 90 deg; joints [18.339, -57.216, 111.169, -157.708, 56.044, 90.139]
  MoveL 746 to (119.22, -33.72, 2.44) mm, rotated rx 90 ry -73.52 rz 90 deg; joints [18.183, -58.267, 110.936, -157.555, 54.821, 93.094]
  MoveL 747 to (120.05, -34.47, 2.68) mm, rotated rx 90 ry -70.08 rz 90 deg; joints [17.977, -59.301, 110.702, -157.453, 53.601, 96.085]
  MoveL 748 to (120.88, -35.2, 2.98) mm, rotated rx 90 ry -66.63 rz 90 deg; joints [17.72, -60.314, 110.468, -157.404, 52.387, 99.116]
  MoveL 749 to (121.71, -35.91, 3.31) mm, rotated rx 90 ry -63.19 rz 90 deg; joints [17.413, -61.304, 110.236, -157.412, 51.181, 102.196]
  MoveL 750 to (122.54, -36.6, 3.69) mm, rotated rx 90 ry -59.74 rz 90 deg; joints [17.058, -62.268, 110.005, -157.481, 49.988, 105.33]
  MoveL 751 to (123.49, -37.13, 4.01) mm, rotated rx 90 ry -57 rz 90 deg; joints [16.736, -63, 109.799, -157.583, 49.037, 107.869]
  MoveL 752 to (124.44, -37.65, 4.37) mm, rotated rx 90 ry -54.25 rz 90 deg; joints [16.385, -63.712, 109.596, -157.729, 48.099, 110.451]
  MoveL 753 to (125.4, -38.15, 4.75) mm, rotated rx 90 ry -51.51 rz 90 deg; joints [16.003, -64.402, 109.397, -157.92, 47.174, 113.078]
  MoveL 754 to (126.35, -38.63, 5.15) mm, rotated rx 90 ry -48.76 rz 90 deg; joints [15.593, -65.069, 109.201, -158.159, 46.265, 115.753]
  MoveL 755 to (127.3, -39.1, 5.58) mm, rotated rx 90 ry -46.01 rz 90 deg; joints [15.155, -65.711, 109.011, -158.449, 45.374, 118.48]
  MoveL 756 to (128.2, -39.35, 5.83) mm, rotated rx 90 ry -44.43 rz 90 deg; joints [14.887, -66.05, 108.874, -158.641, 44.86, 120.073]
  MoveL 757 to (129.1, -39.6, 6.09) mm, rotated rx 90 ry -42.85 rz 90 deg; joints [14.61, -66.38, 108.74, -158.851, 44.354, 121.685]
  MoveL 758 to (130, -39.85, 6.36) mm, rotated rx 90 ry -41.27 rz 90 deg; joints [14.324, -66.701, 108.608, -159.079, 43.855, 123.316]
  MoveL 759 to (130.9, -40.08, 6.63) mm, rotated rx 90 ry -39.69 rz 90 deg; joints [14.029, -67.013, 108.478, -159.326, 43.364, 124.968]
  MoveL 760 to (131.79, -40.31, 6.91) mm, rotated rx 90 ry -38.11 rz 90 deg; joints [13.727, -67.314, 108.35, -159.592, 42.882, 126.64]
  MoveL 761 to (132.69, -40.53, 7.2) mm, rotated rx 90 ry -36.53 rz 90 deg; joints [13.416, -67.607, 108.225, -159.878, 42.409, 128.334]
  MoveL 762 to (133.65, -40.65, 7.37) mm, rotated rx 90 ry -35.62 rz 90 deg; joints [13.23, -67.744, 108.117, -160.052, 42.131, 129.311]
  MoveL 763 to (134.61, -40.77, 7.54) mm, rotated rx 90 ry -34.72 rz 90 deg; joints [13.042, -67.878, 108.011, -160.233, 41.856, 130.296]
  MoveL 764 to (135.57, -40.88, 7.71) mm, rotated rx 90 ry -33.81 rz 90 deg; joints [12.851, -68.008, 107.905, -160.42, 41.584, 131.288]
  MoveL 765 to (136.53, -41, 7.88) mm, rotated rx 90 ry -32.91 rz 90 deg; joints [12.658, -68.135, 107.8, -160.615, 41.316, 132.287]
  MoveL 766 to (137.49, -41.11, 8.06) mm, rotated rx 90 ry -32 rz 90 deg; joints [12.463, -68.258, 107.696, -160.815, 41.052, 133.294]
  MoveL 767 to (138.45, -41.22, 8.23) mm, rotated rx 90 ry -31.1 rz 90 deg; joints [12.266, -68.378, 107.593, -161.023, 40.792, 134.308]
  MoveL 768 to (139.43, -41.23, 8.26) mm, rotated rx 90 ry -30.99 rz 90 deg; joints [12.234, -68.342, 107.509, -161.051, 40.738, 134.428]
  MoveL 769 to (140.41, -41.24, 8.28) mm, rotated rx 90 ry -30.88 rz 90 deg; joints [12.203, -68.306, 107.426, -161.08, 40.685, 134.549]
  MoveL 770 to (141.38, -41.26, 8.3) mm, rotated rx 90 ry -30.77 rz 90 deg; joints [12.172, -68.27, 107.342, -161.109, 40.632, 134.67]
  MoveL 771 to (142.36, -41.27, 8.32) mm, rotated rx 90 ry -30.66 rz 90 deg; joints [12.14, -68.234, 107.258, -161.137, 40.579, 134.789]
  MoveL 772 to (143.34, -41.28, 8.34) mm, rotated rx 90 ry -30.55 rz 90 deg; joints [12.109, -68.198, 107.174, -161.166, 40.525, 134.91]
  MoveL 773 to (144.31, -41.29, 8.36) mm, rotated rx 90 ry -30.45 rz 90 deg; joints [12.078, -68.162, 107.09, -161.195, 40.472, 135.031]
  MoveL 774 to (145.26, -41.2, 8.2) mm, rotated rx 90 ry -31.28 rz 90 deg; joints [12.245, -67.948, 107.032, -161.004, 40.662, 134.081]
  MoveL 775 to (146.21, -41.09, 8.03) mm, rotated rx 90 ry -32.12 rz 90 deg; joints [12.411, -67.731, 106.974, -160.819, 40.855, 133.136]
  MoveL 776 to (147.16, -40.99, 7.87) mm, rotated rx 90 ry -32.96 rz 90 deg; joints [12.574, -67.511, 106.917, -160.64, 41.05, 132.197]
  MoveL 777 to (148.1, -40.89, 7.71) mm, rotated rx 90 ry -33.8 rz 90 deg; joints [12.735, -67.29, 106.861, -160.467, 41.247, 131.265]
  MoveL 778 to (149.05, -40.78, 7.55) mm, rotated rx 90 ry -34.64 rz 90 deg; joints [12.893, -67.065, 106.805, -160.3, 41.447, 130.338]
  MoveL 779 to (150, -40.67, 7.4) mm, rotated rx 90 ry -35.48 rz 90 deg; joints [13.049, -66.838, 106.75, -160.139, 41.65, 129.418]
  MoveL 780 to (150, -41.19, 8.19) mm, rotated rx 90 ry -31.33 rz 90 deg; joints [12.213, -67.664, 106.636, -161.009, 40.548, 134.017]
  MoveL 781 to (150, -41.65, 9.02) mm, rotated rx 90 ry -27.18 rz 90 deg; joints [11.326, -68.422, 106.542, -162.024, 39.521, 138.77]
  MoveL 782 to (150, -42.06, 9.88) mm, rotated rx 90 ry -23.03 rz 90 deg; joints [10.391, -69.108, 106.471, -163.186, 38.577, 143.681]
  MoveL 783 to (150, -42.4, 10.76) mm, rotated rx 90 ry -18.88 rz 90 deg; joints [9.414, -69.72, 106.423, -164.496, 37.726, 148.747]
  MoveL 784 to (150, -42.67, 11.67) mm, rotated rx 90 ry -14.73 rz 90 deg; joints [8.399, -70.253, 106.401, -165.947, 36.98, 153.963]
  MoveL 785 to (150, -42.88, 12.6) mm, rotated rx 90 ry -10.58 rz 90 deg; joints [7.352, -70.708, 106.406, -167.532, 36.349, 159.323]
  MoveL 786 to (150, -43.02, 13.53) mm, rotated rx 90 ry -6.43 rz 90 deg; joints [6.278, -71.079, 106.438, -169.237, 35.84, 164.81]
  MoveL 787 to (150, -43.09, 14.48) mm, rotated rx 90 ry -2.28 rz 90 deg; joints [5.184, -71.367, 106.499, -171.041, 35.464, 170.403]
  MoveL 788 to (150, -43.1, 15.45) mm, rotated rx 90 ry 0 rz 90 deg; joints [4.557, -71.491, 106.548, -172.099, 35.314, 173.539]
  MoveL 789 to (150, -43.1, 16.45) mm, rotated rx 90 ry 0 rz 90 deg; joints [4.516, -71.496, 106.555, -172.171, 35.311, 173.598]
  MoveL 790 to (150, -43.1, 17.44) mm, rotated rx 90 ry 0 rz 90 deg; joints [4.475, -71.501, 106.561, -172.242, 35.308, 173.656]
  MoveL 791 to (150, -43.1, 18.44) mm, rotated rx 90 ry 0 rz 90 deg; joints [4.433, -71.506, 106.568, -172.314, 35.306, 173.715]
  MoveL 792 to (150, -43.1, 19.43) mm, rotated rx 90 ry 0 rz 90 deg; joints [4.392, -71.51, 106.574, -172.385, 35.303, 173.773]
  MoveL 793 to (150, -43.1, 20.43) mm, rotated rx 90 ry 0 rz 90 deg; joints [4.35, -71.515, 106.58, -172.457, 35.3, 173.832]
  MoveL 794 to (150, -43.1, 21.42) mm, rotated rx 90 ry 0 rz 90 deg; joints [4.309, -71.52, 106.587, -172.528, 35.297, 173.89]
  MoveL 795 to (150, -43.1, 22.42) mm, rotated rx 90 ry 0 rz 90 deg; joints [4.268, -71.524, 106.593, -172.6, 35.294, 173.949]
  MoveL 796 to (150, -43.1, 23.42) mm, rotated rx 90 ry 0 rz 90 deg; joints [4.226, -71.529, 106.599, -172.672, 35.292, 174.008]
  MoveL 797 to (150, -43.1, 24.41) mm, rotated rx 90 ry 0 rz 90 deg; joints [4.185, -71.533, 106.605, -172.743, 35.289, 174.066]
  MoveL 798 to (150, -43.1, 25.41) mm, rotated rx 90 ry 0 rz 90 deg; joints [4.143, -71.538, 106.611, -172.815, 35.286, 174.125]
  MoveL 799 to (150, -43.1, 26.4) mm, rotated rx 90 ry 0 rz 90 deg; joints [4.102, -71.542, 106.617, -172.886, 35.284, 174.183]
  MoveL 800 to (150, -43.1, 27.4) mm, rotated rx 90 ry 0 rz 90 deg; joints [4.06, -71.546, 106.623, -172.958, 35.281, 174.242]
  MoveL 801 to (150, -43.1, 28.39) mm, rotated rx 90 ry 0 rz 90 deg; joints [4.019, -71.551, 106.629, -173.03, 35.278, 174.3]
  MoveL 802 to (150, -43.1, 29.39) mm, rotated rx 90 ry 0 rz 90 deg; joints [3.978, -71.555, 106.635, -173.101, 35.276, 174.359]
  MoveL 803 to (150, -43.1, 30.39) mm, rotated rx 90 ry 0 rz 90 deg; joints [3.936, -71.559, 106.64, -173.173, 35.273, 174.418]
  MoveL 804 to (150, -43.1, 31.38) mm, rotated rx 90 ry 0 rz 90 deg; joints [3.895, -71.563, 106.646, -173.245, 35.271, 174.476]
  MoveL 805 to (150, -43.1, 32.38) mm, rotated rx 90 ry 0 rz 90 deg; joints [3.853, -71.568, 106.652, -173.316, 35.268, 174.535]
  MoveL 806 to (150, -43.1, 33.37) mm, rotated rx 90 ry 0 rz 90 deg; joints [3.812, -71.572, 106.657, -173.388, 35.266, 174.594]
  MoveL 807 to (150, -43.1, 34.37) mm, rotated rx 90 ry 0 rz 90 deg; joints [3.77, -71.576, 106.663, -173.46, 35.263, 174.652]
  MoveL 808 to (150, -43.1, 35.37) mm, rotated rx 90 ry 0 rz 90 deg; joints [3.729, -71.58, 106.668, -173.532, 35.261, 174.711]
  MoveL 809 to (150, -43.1, 36.36) mm, rotated rx 90 ry 0 rz 90 deg; joints [3.687, -71.584, 106.674, -173.603, 35.258, 174.77]
  MoveL 810 to (150, -43.1, 37.36) mm, rotated rx 90 ry 0 rz 90 deg; joints [3.646, -71.588, 106.679, -173.675, 35.256, 174.828]
  MoveL 811 to (150, -43.1, 38.35) mm, rotated rx 90 ry 0 rz 90 deg; joints [3.604, -71.591, 106.684, -173.747, 35.254, 174.887]
  MoveL 812 to (150, -43.1, 39.35) mm, rotated rx 90 ry 0 rz 90 deg; joints [3.563, -71.595, 106.689, -173.819, 35.251, 174.946]
  MoveL 813 to (150, -43.1, 40.34) mm, rotated rx 90 ry 0 rz 90 deg; joints [3.521, -71.599, 106.694, -173.891, 35.249, 175.004]
  MoveL 814 to (150, -43.1, 41.34) mm, rotated rx 90 ry 0 rz 90 deg; joints [3.48, -71.603, 106.7, -173.962, 35.247, 175.063]
  MoveL 815 to (150, -43.1, 42.34) mm, rotated rx 90 ry 0 rz 90 deg; joints [3.438, -71.607, 106.705, -174.034, 35.244, 175.122]
  MoveL 816 to (143.45, -43.1, 34.64) mm, rotated rx 90 ry 0 rz 90 deg; joints [3.777, -71.979, 107.208, -173.471, 35.405, 174.671]
  MoveL 817 to (140.08, -43.1, 30.93) mm, rotated rx 90 ry 0 rz 90 deg; joints [3.942, -72.17, 107.465, -173.199, 35.487, 174.453]
  MoveL 818 to (139.31, -43.1, 29.9) mm, rotated rx 90 ry 0 rz 90 deg; joints [3.988, -72.213, 107.523, -173.123, 35.506, 174.393]
  MoveL 819 to (138.55, -43.1, 28.85) mm, rotated rx 90 ry 0 rz 90 deg; joints [4.034, -72.255, 107.58, -173.047, 35.525, 174.332]
  MoveL 820 to (137.52, -43.1, 28.32) mm, rotated rx 90 ry 0 rz 90 deg; joints [4.059, -72.316, 107.661, -173.007, 35.548, 174.301]
  MoveL 821 to (136.22, -43.1, 28.33) mm, rotated rx 90 ry 0 rz 90 deg; joints [4.062, -72.395, 107.768, -173.006, 35.575, 174.302]
  MoveL 822 to (129.47, -43.1, 28.85) mm, rotated rx 90 ry 0 rz 90 deg; joints [4.061, -72.812, 108.325, -173.032, 35.715, 174.333]
  MoveL 823 to (122.87, -43.1, 29.88) mm, rotated rx 90 ry 0 rz 90 deg; joints [4.037, -73.221, 108.87, -173.096, 35.847, 174.394]
  MoveL 824 to (116.19, -43.1, 31.26) mm, rotated rx 90 ry 0 rz 90 deg; joints [3.998, -73.637, 109.421, -173.183, 35.976, 174.475]
  MoveL 825 to (106.18, -43.1, 32.79) mm, rotated rx 90 ry 0 rz 90 deg; joints [3.962, -74.258, 110.237, -173.275, 36.166, 174.563]
  MoveL 826 to (96.14, -43.1, 33.56) mm, rotated rx 90 ry 0 rz 90 deg; joints [3.959, -74.879, 111.044, -173.311, 36.352, 174.604]
  MoveL 827 to (86.07, -43.1, 34.2) mm, rotated rx 90 ry 0 rz 90 deg; joints [3.962, -75.501, 111.848, -173.335, 36.532, 174.636]
  MoveL 828 to (75.98, -43.1, 34.65) mm, rotated rx 90 ry 0 rz 90 deg; joints [3.973, -76.125, 112.646, -173.344, 36.707, 174.655]
  MoveL 829 to (71.53, -43.1, 34.01) mm, rotated rx 90 ry 0 rz 90 deg; joints [4.015, -76.397, 112.991, -173.286, 36.784, 174.614]
  MoveL 830 to (67.42, -43.1, 32.19) mm, rotated rx 90 ry 0 rz 90 deg; joints [4.108, -76.643, 113.303, -173.141, 36.857, 174.503]
  MoveL 831 to (64.23, -43.1, 29.07) mm, rotated rx 90 ry 0 rz 90 deg; joints [4.257, -76.825, 113.533, -172.902, 36.919, 174.315]
  MoveL 832 to (62.23, -43.1, 24.95) mm, rotated rx 90 ry 0 rz 90 deg; joints [4.446, -76.929, 113.664, -172.593, 36.965, 174.07]
  MoveL 833 to (61.36, -43.1, 20.36) mm, rotated rx 90 ry 0 rz 90 deg; joints [4.653, -76.961, 113.704, -172.253, 36.995, 173.799]
  MoveL 834 to (61.51, -43.1, 15.75) mm, rotated rx 90 ry 0 rz 90 deg; joints [4.857, -76.928, 113.662, -171.914, 37.009, 173.527]
  MoveL 835 to (61.7, -43.1, 14.88) mm, rotated rx 90 ry -0.54 rz 90 deg; joints [5.043, -76.884, 113.631, -171.61, 37.044, 172.75]
  MoveL 836 to (61.89, -43.07, 14.04) mm, rotated rx 90 ry -4.21 rz 90 deg; joints [6.083, -76.636, 113.553, -169.939, 37.345, 167.762]
  MoveL 837 to (62.08, -42.98, 13.2) mm, rotated rx 90 ry -7.88 rz 90 deg; joints [7.109, -76.316, 113.499, -168.341, 37.76, 162.852]
  MoveL 838 to (62.27, -42.83, 12.38) mm, rotated rx 90 ry -11.56 rz 90 deg; joints [8.114, -75.925, 113.467, -166.831, 38.282, 158.035]
  MoveL 839 to (62.46, -42.64, 11.56) mm, rotated rx 90 ry -15.23 rz 90 deg; joints [9.096, -75.466, 113.459, -165.421, 38.906, 153.328]
  MoveL 840 to (62.75, -42.4, 10.78) mm, rotated rx 90 ry -18.77 rz 90 deg; joints [10.013, -74.953, 113.462, -164.168, 39.593, 148.905]
  MoveL 841 to (63.05, -42.12, 10.03) mm, rotated rx 90 ry -22.31 rz 90 deg; joints [10.901, -74.38, 113.485, -163.021, 40.361, 144.597]
  MoveL 842 to (63.35, -41.79, 9.29) mm, rotated rx 90 ry -25.84 rz 90 deg; joints [11.755, -73.747, 113.526, -161.984, 41.201, 140.406]
  MoveL 843 to (63.65, -41.41, 8.57) mm, rotated rx 90 ry -29.38 rz 90 deg; joints [12.573, -73.059, 113.585, -161.056, 42.108, 136.333]
  MoveL 844 to (63.95, -41, 7.88) mm, rotated rx 90 ry -32.92 rz 90 deg; joints [13.351, -72.315, 113.659, -160.237, 43.074, 132.375]
  MoveL 845 to (64.26, -40.53, 7.21) mm, rotated rx 90 ry -36.52 rz 90 deg; joints [14.1, -71.506, 113.748, -159.513, 44.11, 128.468]
  MoveL 846 to (64.58, -40.02, 6.56) mm, rotated rx 90 ry -40.11 rz 90 deg; joints [14.803, -70.645, 113.85, -158.893, 45.193, 124.671]
  MoveL 847 to (64.89, -39.47, 5.95) mm, rotated rx 90 ry -43.71 rz 90 deg; joints [15.458, -69.735, 113.964, -158.374, 46.319, 120.98]
  MoveL 848 to (65.21, -38.88, 5.37) mm, rotated rx 90 ry -47.3 rz 90 deg; joints [16.064, -68.779, 114.088, -157.949, 47.481, 117.387]
  MoveL 849 to (65.53, -38.26, 4.83) mm, rotated rx 90 ry -50.9 rz 90 deg; joints [16.619, -67.781, 114.221, -157.614, 48.674, 113.886]
  MoveL 850 to (65.76, -37.59, 4.32) mm, rotated rx 90 ry -54.58 rz 90 deg; joints [17.134, -66.722, 114.371, -157.356, 49.926, 110.385]
  MoveL 851 to (66, -36.89, 3.86) mm, rotated rx 90 ry -58.27 rz 90 deg; joints [17.593, -65.624, 114.527, -157.181, 51.2, 106.962]
  MoveL 852 to (66.23, -36.16, 3.44) mm, rotated rx 90 ry -61.95 rz 90 deg; joints [17.994, -64.491, 114.686, -157.082, 52.493, 103.611]
  MoveL 853 to (66.47, -35.4, 3.07) mm, rotated rx 90 ry -65.64 rz 90 deg; joints [18.337, -63.327, 114.849, -157.054, 53.798, 100.323]
  MoveL 854 to (66.7, -34.62, 2.74) mm, rotated rx 90 ry -69.32 rz 90 deg; joints [18.62, -62.136, 115.012, -157.092, 55.113, 97.09]
  MoveL 855 to (66.96, -33.83, 2.47) mm, rotated rx 90 ry -72.98 rz 90 deg; joints [18.842, -60.931, 115.172, -157.192, 56.423, 93.928]
  MoveL 856 to (67.21, -33.03, 2.25) mm, rotated rx 90 ry -76.64 rz 90 deg; joints [19.005, -59.706, 115.33, -157.349, 57.735, 90.805]
  MoveL 857 to (67.47, -32.21, 2.09) mm, rotated rx 90 ry -80.29 rz 90 deg; joints [19.108, -58.467, 115.486, -157.559, 59.045, 87.715]
  MoveL 858 to (67.72, -31.38, 1.97) mm, rotated rx 90 ry -83.95 rz 90 deg; joints [19.152, -57.218, 115.638, -157.821, 60.35, 84.649]
  MoveL 859 to (68.18, -30.66, 1.92) mm, rotated rx 90 ry -87.11 rz 90 deg; joints [19.138, -56.122, 115.746, -158.088, 61.463, 82.011]
  MoveL 860 to (68.65, -29.93, 1.9) mm, rotated rx 0 ry -90 rz 180 deg; joints [19.086, -55.115, 115.839, -158.364, 62.475, 79.612]
  MoveL 861 to (69.11, -29.18, 1.9) mm, rotated rx 0 ry -90 rz 180 deg; joints [19.079, -55.055, 115.805, -158.376, 62.498, 79.627]
  MoveL 862 to (69.58, -28.42, 1.9) mm, rotated rx 0 ry -90 rz 180 deg; joints [19.073, -54.994, 115.771, -158.388, 62.522, 79.641]
  MoveL 863 to (72.19, -25.91, 1.9) mm, rotated rx 0 ry -90 rz 180 deg; joints [19.037, -54.749, 115.57, -158.436, 62.557, 79.678]
  MoveL 864 to (74.99, -23.64, 1.9) mm, rotated rx 0 ry -90 rz 180 deg; joints [18.999, -54.509, 115.354, -158.483, 62.571, 79.707]
  MoveL 865 to (77.89, -21.53, 1.9) mm, rotated rx 0 ry -90 rz 180 deg; joints [18.959, -54.274, 115.127, -158.528, 62.572, 79.73]
  MoveL 866 to (86.56, -15.59, 1.9) mm, rotated rx 0 ry -90 rz 180 deg; joints [18.842, -53.591, 114.443, -158.657, 62.55, 79.789]
  MoveL 867 to (95.34, -9.78, 1.9) mm, rotated rx 0 ry -90 rz 180 deg; joints [18.725, -52.914, 113.742, -158.783, 62.508, 79.84]
  MoveL 868 to (100.49, -6.86, 1.9) mm, rotated rx 0 ry -90 rz 180 deg; joints [18.658, -52.543, 113.327, -158.85, 62.455, 79.857]
  MoveL 869 to (105.92, -4.55, 1.9) mm, rotated rx 0 ry -90 rz 180 deg; joints [18.586, -52.194, 112.885, -158.912, 62.355, 79.855]
  MoveL 870 to (109.55, -3.6, 1.9) mm, rotated rx 0 ry -90 rz 180 deg; joints [18.539, -51.992, 112.587, -158.946, 62.257, 79.841]
  MoveL 871 to (113.24, -2.81, 1.9) mm, rotated rx 0 ry -90 rz 180 deg; joints [18.491, -51.796, 112.283, -158.979, 62.148, 79.822]
  MoveL 872 to (116.81, -1.76, 1.9) mm, rotated rx 0 ry -90 rz 180 deg; joints [18.445, -51.591, 111.988, -159.013, 62.056, 79.809]
  MoveL 873 to (120.13, 0, 1.9) mm, rotated rx 0 ry -90 rz 180 deg; joints [18.403, -51.36, 111.715, -159.053, 62.01, 79.815]
  MoveL 874 to (89.24, 0, 1.9) mm, rotated rx 0 ry -90 rz 180 deg; joints [18.807, -52.635, 114.264, -158.841, 63.268, 80.124]
  MoveL 875 to (82.11, -4.36, 1.9) mm, rotated rx 0 ry -90 rz 180 deg; joints [18.902, -53.165, 114.835, -158.743, 63.323, 80.093]
  MoveL 876 to (75.14, -9.38, 1.9) mm, rotated rx 0 ry -90 rz 180 deg; joints [18.997, -53.725, 115.389, -158.638, 63.333, 80.044]
  MoveL 877 to (68.48, -14.73, 1.9) mm, rotated rx 0 ry -90 rz 180 deg; joints [19.088, -54.292, 115.911, -158.529, 63.307, 79.98]
  MoveL 878 to (63.8, -18.78, 1.9) mm, rotated rx 0 ry -90 rz 180 deg; joints [19.152, -54.708, 116.274, -158.448, 63.269, 79.927]
  MoveL 879 to (59.46, -22.76, 1.9) mm, rotated rx 0 ry -90 rz 180 deg; joints [19.213, -55.106, 116.607, -158.37, 63.22, 79.87]
  MoveL 880 to (55.29, -27.11, 1.9) mm, rotated rx 0 ry -90 rz 180 deg; joints [19.271, -55.519, 116.924, -158.288, 63.141, 79.802]
  MoveL 881 to (53.14, -29.73, 1.9) mm, rotated rx 0 ry -90 rz 180 deg; joints [19.301, -55.752, 117.084, -158.241, 63.079, 79.756]
  MoveL 882 to (52.59, -30.45, 1.91) mm, rotated rx 90 ry -88.05 rz 90 deg; joints [19.344, -56.464, 117.039, -158.048, 62.384, 81.367]
  MoveL 883 to (52.04, -31.15, 1.95) mm, rotated rx 90 ry -84.95 rz 90 deg; joints [19.373, -57.557, 116.94, -157.776, 61.285, 83.939]
  MoveL 884 to (51.36, -31.44, 1.98) mm, rotated rx 90 ry -83.7 rz 90 deg; joints [19.379, -58.019, 116.936, -157.672, 60.854, 84.987]
  MoveL 885 to (50.68, -31.72, 2.01) mm, rotated rx 90 ry -82.45 rz 90 deg; joints [19.377, -58.481, 116.931, -157.573, 60.422, 86.038]
  MoveL 886 to (50, -32.01, 2.06) mm, rotated rx 90 ry -81.19 rz 90 deg; joints [19.369, -58.943, 116.925, -157.48, 59.988, 87.091]
  MoveL 887 to (49.35, -31.89, 2.04) mm, rotated rx 90 ry -81.71 rz 90 deg; joints [19.387, -58.794, 117.002, -157.51, 60.201, 86.663]
  MoveL 888 to (48.7, -31.77, 2.02) mm, rotated rx 90 ry -82.23 rz 90 deg; joints [19.403, -58.644, 117.078, -157.541, 60.413, 86.235]
  MoveL 889 to (48.09, -31.09, 1.95) mm, rotated rx 90 ry -85.2 rz 90 deg; joints [19.429, -57.643, 117.267, -157.763, 61.518, 83.766]
  MoveL 890 to (47.47, -30.42, 1.91) mm, rotated rx 90 ry -88.17 rz 90 deg; joints [19.415, -56.637, 117.452, -158.017, 62.619, 81.308]
  MoveL 891 to (46.86, -29.73, 1.9) mm, rotated rx 0 ry -90 rz 180 deg; joints [19.389, -56.012, 117.584, -158.188, 63.317, 79.812]
  MoveL 892 to (44.71, -27.11, 1.9) mm, rotated rx 0 ry -90 rz 180 deg; joints [19.42, -55.956, 117.766, -158.199, 63.543, 79.896]
  MoveL 893 to (40.54, -22.76, 1.9) mm, rotated rx 0 ry -90 rz 180 deg; joints [19.479, -55.885, 118.115, -158.211, 63.944, 80.041]
  MoveL 894 to (36.2, -18.78, 1.9) mm, rotated rx 0 ry -90 rz 180 deg; joints [19.542, -55.839, 118.474, -158.215, 64.33, 80.178]
  MoveL 895 to (31.52, -14.73, 1.9) mm, rotated rx 0 ry -90 rz 180 deg; joints [19.609, -55.798, 118.857, -158.217, 64.735, 80.32]
  MoveL 896 to (24.86, -9.38, 1.9) mm, rotated rx 0 ry -90 rz 180 deg; joints [19.706, -55.759, 119.397, -158.211, 65.289, 80.513]
  MoveL 897 to (17.89, -4.36, 1.9) mm, rotated rx 0 ry -90 rz 180 deg; joints [19.808, -55.746, 119.956, -158.197, 65.837, 80.701]
  MoveL 898 to (10.76, 0, 1.9) mm, rotated rx 0 ry -90 rz 180 deg; joints [19.914, -55.771, 120.522, -158.172, 66.356, 80.874]
  MoveL 899 to (29.57, 0, 1.9) mm, rotated rx 0 ry -90 rz 180 deg; joints [19.637, -55.033, 119.049, -158.35, 65.63, 80.698]
  MoveL 900 to (32.44, -3.98, 1.9) mm, rotated rx 0 ry -90 rz 180 deg; joints [19.596, -55.148, 118.814, -158.336, 65.297, 80.575]
  MoveL 901 to (36.09, -7.89, 1.9) mm, rotated rx 0 ry -90 rz 180 deg; joints [19.543, -55.225, 118.516, -158.329, 64.94, 80.446]
  MoveL 902 to (39.95, -11.79, 1.9) mm, rotated rx 0 ry -90 rz 180 deg; joints [19.488, -55.291, 118.2, -158.323, 64.575, 80.315]
  MoveL 903 to (42.66, -14.76, 1.9) mm, rotated rx 0 ry -90 rz 180 deg; joints [19.449, -55.349, 117.975, -158.315, 64.306, 80.218]
  MoveL 904 to (44.97, -17.81, 1.9) mm, rotated rx 0 ry -90 rz 180 deg; joints [19.416, -55.427, 117.782, -158.302, 64.049, 80.123]
  MoveL 905 to (46.69, -20.99, 1.9) mm, rotated rx 0 ry -90 rz 180 deg; joints [19.392, -55.534, 117.634, -158.283, 63.808, 80.029]
  MoveL 906 to (47.76, -22.83, 1.9) mm, rotated rx 0 ry -90 rz 180 deg; joints [19.377, -55.593, 117.542, -158.272, 63.665, 79.974]
  MoveL 907 to (48.52, -23.66, 1.9) mm, rotated rx 0 ry -90 rz 180 deg; joints [19.366, -55.608, 117.478, -158.269, 63.59, 79.947]
  MoveL 908 to (50, -24, 1.9) mm, rotated rx 0 ry -90 rz 180 deg; joints [19.345, -55.565, 117.359, -158.278, 63.515, 79.925]
  MoveL 909 to (51.48, -23.66, 1.9) mm, rotated rx 0 ry -90 rz 180 deg; joints [19.324, -55.486, 117.242, -158.294, 63.477, 79.92]
  MoveL 910 to (52.24, -22.83, 1.9) mm, rotated rx 0 ry -90 rz 180 deg; joints [19.314, -55.408, 117.184, -158.31, 63.493, 79.934]
  MoveL 911 to (53.31, -20.99, 1.9) mm, rotated rx 0 ry -90 rz 180 deg; joints [19.298, -55.262, 117.106, -158.339, 63.554, 79.969]
  MoveL 912 to (54.11, -19.37, 1.9) mm, rotated rx 0 ry -90 rz 180 deg; joints [19.287, -55.139, 117.048, -158.363, 63.612, 80.001]
  MoveL 913 to (55.03, -17.81, 1.9) mm, rotated rx 0 ry -90 rz 180 deg; joints [19.274, -55.015, 116.98, -158.388, 63.662, 80.031]
  MoveL 914 to (57.34, -14.76, 1.9) mm, rotated rx 0 ry -90 rz 180 deg; joints [19.242, -54.751, 116.806, -158.439, 63.739, 80.083]
  MoveL 915 to (60.05, -11.79, 1.9) mm, rotated rx 0 ry -90 rz 180 deg; joints [19.204, -54.476, 116.597, -158.493, 63.795, 80.129]
  MoveL 916 to (63.91, -7.89, 1.9) mm, rotated rx 0 ry -90 rz 180 deg; joints [19.151, -54.102, 116.298, -158.565, 63.856, 80.185]
  MoveL 917 to (67.56, -3.98, 1.9) mm, rotated rx 0 ry -90 rz 180 deg; joints [19.101, -53.737, 116.014, -158.635, 63.922, 80.242]
  MoveL 918 to (70.43, 0, 1.9) mm, rotated rx 0 ry -90 rz 180 deg; joints [19.061, -53.4, 115.791, -158.698, 64.022, 80.308]
  MoveL 919 to (70.43, 0, -43.1) mm, rotated rx 0 ry -90 rz 180 deg; joints [20.826, -52.741, 114.474, -156.641, 63.728, 79.177]
  END
